(* PLC project Vn_ld_falling_contact, Beckhoff Automation GmbH TwinCAT PLC Control 3.5.13.21 *)
(* stored: creationDateTime 1970-01-01T00:00:00 *)

PROGRAM Vn_ld_falling_contact
  VAR  (* added by the conversion: wires and edge detectors of the diagram *)
    F_TRIG1 : F_TRIG;
  END_VAR

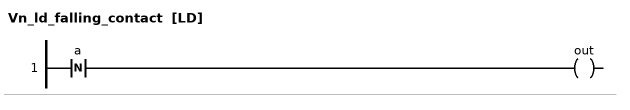
(* LD diagram, written out as Structured Text *)
F_TRIG1(CLK := a);
out := F_TRIG1.Q;
END_PROGRAM
